(* IEC 61131-3 sources: ZPLC/packages/zplc-ide/projects/il_typed_steps_starter/src, 1 file *)

(* ---- TypedSteps.il ---- *)
PROGRAM TypedSteps
VAR_INPUT
    Step AT %I0.0 : BOOL;
    Reset AT %I0.1 : BOOL;
END_VAR
VAR_OUTPUT
    Low AT %Q0.0 : BOOL;
    Exact AT %Q0.1 : BOOL;
    High AT %Q0.2 : BOOL;
END_VAR
VAR
    Total : INT := 0;
    StepWas : BOOL := FALSE;
END_VAR

(* Exercise: add 5 to Total on each rising edge of Step, and clear Total while Reset is TRUE. *)
        LD    Step
        ST    StepWas
        LD    Total
        LT    10
        ST    Low
        LD    Total
        EQ    10
        ST    Exact
        LD    Total
        GT    10
        ST    High
END_PROGRAM
